(* PLC project station_cds.project, CODESYS CODESYS V3.5 SP22 Patch 1 *)
(* stored: creationDateTime 2026-11-25T17:27:32.309646, modificationDateTime 2026-11-25T17:27:31.3827148 *)

FUNCTION_BLOCK FB_HandleStation
  VAR_INPUT
    CycleTime : REAL := 0.002;  (* s *)
    SafetyOk : BOOL;
    DriveOk : BOOL;
    AckFault : BOOL;
    StartEnable : BOOL;  (* release from the line *)
    PartPresent : BOOL;
    SensLH : BOOL;  (* variant sensor that only an LH unit covers *)
    SensRH : BOOL;  (* variant sensor that only an RH unit covers *)
    VariantLH : BOOL;  (* recipe: TRUE = LH units are being built *)
    ClampClosed : BOOL;
    ClampOpen : BOOL;
    RejectChute : BOOL;  (* light barrier in the reject chute *)
    Pos : REAL;  (* mm, axis position, 0 = home *)
    Force : REAL;  (* N, load cell *)
    VPull : REAL := 50.0;  (* mm/s *)
    VHome : REAL := 150.0;  (* mm/s *)
    FTouch : REAL := 1.5;  (* N *)
    FRev : REAL := 40.0;  (* N *)
    FAbsMax : REAL := 60.0;  (* N, protects the painted part *)
    XMax : REAL := 38.0;  (* mm *)
    TouchLo : REAL := 3.0;  (* mm, window of the touch position *)
    TouchHi : REAL := 7.0;
    Compliance : REAL := 0.025;  (* mm/N, rig deflection taken out of the travel *)
    TareTol : REAL := 0.5;  (* N *)
    TPresent : REAL := 0.1;  (* s *)
    TClampMax : REAL := 1.0;  (* s *)
    TRejectWarn : REAL := 30.0;  (* s *)
    MaxConsecNok : INT := 3;
  END_VAR
  VAR_IN_OUT
    Rcp : ST_EvalRecipe;  (* evaluation recipe, copied into Eval at every tare *)
  END_VAR
  VAR_OUTPUT
    QClamp : BOOL;
    QDriveEnable : BOOL;
    QVel : REAL;  (* mm/s, positive = pull *)
    QLampOk : BOOL;
    QLampNok : BOOL;
    QCallOperator : BOOL;
    State : INT;
    Verdict : INT;  (* 0 none, 1 OK, 2 NOK *)
    NokCode : INT;
    FaultCode : INT;
    Locked : BOOL;
    RigCheckRequired : BOOL;  (* too many rejects in a row: run the master part *)
    XTravel : REAL;  (* mm *)
    FNet : REAL;  (* N *)
    TCycle : REAL;  (* s, clamp to verdict of the last part *)
    CntTotal : DINT;
    CntOk : DINT;
    CntNok : DINT;
    CntRejectConfirmed : DINT;
    CntConsecNok : INT;
    CntByCode : ARRAY[0..31] OF DINT;
  END_VAR
  VAR
    Eval : FB_CurveEval;
    sTim : REAL;
    sTCycle : REAL;
    sTare : REAL;
    sTouchPos : REAL;
    sFTouch : REAL;
    sPreNok : INT;
    sPartGone : BOOL;
    sChutePrev : BOOL;
    sInTest : BOOL;
    sWasLocked : BOOL;
    sState : INT;
    sRigCheckRequired : BOOL;
    sCntTotal : DINT;
    sCntOk : DINT;
    sCntNok : DINT;
    sCntRejectConfirmed : DINT;
    sCntConsecNok : INT;
    sCntByCode : ARRAY[0..31] OF DINT;
  END_VAR
  VAR_TEMP
    tVariantOk : BOOL;
    tChuteEdge : BOOL;
    tCode : INT;
  END_VAR

                {region "Inputs"}
        FNet := Force - sTare;
        tChuteEdge := RejectChute AND NOT sChutePrev;
        sChutePrev := RejectChute;
        sTim := sTim + CycleTime;
        sTCycle := sTCycle + CycleTime;
        QVel := 0.0;
        // exactly the sensor of the expected hand, and not the other one
        tVariantOk := (VariantLH AND SensLH AND NOT SensRH) OR (NOT VariantLH AND SensRH AND NOT SensLH);
    {endregion}

    {region "Faults"}
        IF sState <> 9 AND (NOT SafetyOk OR NOT DriveOk) THEN
            IF NOT SafetyOk THEN
                FaultCode := 1;
            ELSE
                FaultCode := 2;
            END_IF;
            IF sState <> 10 THEN
                sInTest := sState >= 1 AND sState <= 6;
                sWasLocked := sState = 8;
            END_IF;
            sState := 9;
        END_IF;
    {endregion}

    {region "Sequence"}
        CASE sState OF
            0:  // Idle
                Locked := FALSE;
                IF NOT PartPresent THEN
                    sTim := 0.0;
                    QLampOk := FALSE;
                    QLampNok := FALSE;
                ELSIF sTim >= TPresent AND StartEnable AND ClampOpen AND NOT sRigCheckRequired THEN
                    Verdict := 0;
                    NokCode := 0;
                    sPreNok := 0;
                    sTCycle := 0.0;
                    sTim := 0.0;
                    IF tVariantOk THEN
                        sState := 1;
                    ELSE
                        sPreNok := 20;   // never pull a part of the wrong hand
                        sState := 6;
                    END_IF;
                END_IF;
            1:  // Clamp
                QClamp := TRUE;
                IF ClampClosed THEN
                    sTim := 0.0;
                    sState := 2;
                ELSIF sTim > TClampMax THEN
                    FaultCode := 3;
                    sInTest := TRUE;
                    sState := 9;
                END_IF;
            2:  // Tare
                IF sTim >= 0.05 THEN
                    IF ABS(Force) > TareTol THEN
                        FaultCode := 4;
                        sInTest := TRUE;
                        sState := 9;
                    ELSE
                        sTare := Force;
                        // the recipe of this part (Siemens: written into Eval by the caller)
                        Eval.Mode := Rcp.Mode;
                        Eval.GateX := Rcp.GateX;
                        Eval.Gate2X := Rcp.Gate2X;
                        Eval.PeakXLo := Rcp.PeakXLo;
                        Eval.PeakXHi := Rcp.PeakXHi;
                        Eval.StepSpan := Rcp.StepSpan;
                        Eval.StopF := Rcp.StopF;
                        Eval.G1Lo := Rcp.G1Lo;
                        Eval.G1Hi := Rcp.G1Hi;
                        Eval.MeanLo := Rcp.MeanLo;
                        Eval.MeanHi := Rcp.MeanHi;
                        Eval.HystLo := Rcp.HystLo;
                        Eval.HystHi := Rcp.HystHi;
                        Eval.RetFMin := Rcp.RetFMin;
                        Eval.G2Lo := Rcp.G2Lo;
                        Eval.G2Hi := Rcp.G2Hi;
                        Eval.PeakFLo := Rcp.PeakFLo;
                        Eval.PeakFHi := Rcp.PeakFHi;
                        Eval.PeakXMin := Rcp.PeakXMin;
                        Eval.PeakXMax := Rcp.PeakXMax;
                        Eval.StepLo := Rcp.StepLo;
                        Eval.StopXLo := Rcp.StopXLo;
                        Eval.StopXHi := Rcp.StopXHi;
                        Eval.EnvX0 := Rcp.EnvX0;
                        Eval.EnvDx := Rcp.EnvDx;
                        Eval.EnvN := Rcp.EnvN;
                        Eval.EnvLo := Rcp.EnvLo;
                        Eval.EnvHi := Rcp.EnvHi;
                        Eval(Reset := TRUE, Sample := FALSE, Stroke := 0, X := 0.0, F := 0.0, Finish := FALSE);
                        sState := 3;
                    END_IF;
                END_IF;
            3:  // Approach
                QVel := VPull;
                IF FNet > FTouch THEN
                    sTouchPos := Pos;
                    sFTouch := FNet;
                    IF Pos < TouchLo OR Pos > TouchHi THEN
                        sPreNok := 21;
                        sState := 5;
                    ELSE
                        XTravel := 0.0;
                        Eval(Reset := FALSE, Sample := TRUE, Stroke := 1, X := 0.0, F := FNet, Finish := FALSE);
                        sState := 4;
                    END_IF;
                ELSIF Pos > TouchHi THEN
                    sPreNok := 21;
                    sTouchPos := Pos;
                    sFTouch := 0.0;
                    sState := 5;
                END_IF;
            4:  // Pull
                QVel := VPull;
                XTravel := Pos - sTouchPos - (FNet - sFTouch) * Compliance;
                Eval(Reset := FALSE, Sample := TRUE, Stroke := 1, X := XTravel, F := FNet, Finish := FALSE);
                IF FNet >= FAbsMax THEN
                    sPreNok := 22;
                    sState := 5;
                ELSIF FNet >= FRev THEN
                    sState := 5;
                ELSIF XTravel >= XMax THEN
                    sPreNok := 23;
                    sState := 5;
                END_IF;
            5:  // Return
                XTravel := Pos - sTouchPos - (FNet - sFTouch) * Compliance;
                IF Pos > sTouchPos - 0.5 THEN
                    QVel := -VPull;
                    IF sPreNok = 0 THEN
                        Eval(Reset := FALSE, Sample := TRUE, Stroke := 2, X := XTravel, F := FNet, Finish := FALSE);
                    END_IF;
                ELSIF Pos > 0.05 THEN
                    QVel := -VHome;
                ELSE
                    sState := 6;
                END_IF;
            6:  // Evaluate
                IF sPreNok <> 0 THEN
                    tCode := sPreNok;
                ELSE
                    Eval(Reset := FALSE, Sample := FALSE, Stroke := 0, X := 0.0, F := 0.0, Finish := TRUE);
                    tCode := Eval.NokCode;
                END_IF;
                NokCode := tCode;
                TCycle := sTCycle;
                sCntTotal := sCntTotal + 1;
                sCntByCode[tCode] := sCntByCode[tCode] + 1;
                QClamp := FALSE;
                sTim := 0.0;
                IF tCode = 0 THEN
                    Verdict := 1;
                    sCntOk := sCntOk + 1;
                    sCntConsecNok := 0;
                    QLampOk := TRUE;
                    sState := 7;
                ELSE
                    Verdict := 2;
                    sCntNok := sCntNok + 1;
                    sCntConsecNok := sCntConsecNok + 1;
                    QLampNok := TRUE;
                    sPartGone := FALSE;
                    sState := 8;
                END_IF;
            7:  // UnloadOk
                QClamp := FALSE;
                IF NOT PartPresent AND ClampOpen THEN
                    sTim := 0.0;
                    sState := 0;
                END_IF;
            8:  // RejectLock
                QClamp := FALSE;
                Locked := TRUE;
                IF NOT PartPresent THEN
                    sPartGone := TRUE;
                END_IF;
                QCallOperator := sTim > TRejectWarn OR sRigCheckRequired;
                IF sPartGone AND tChuteEdge THEN
                    sCntRejectConfirmed := sCntRejectConfirmed + 1;
                    sRigCheckRequired := sCntConsecNok >= MaxConsecNok;
                    QCallOperator := sRigCheckRequired;
                    Locked := FALSE;
                    sTim := 0.0;
                    sState := 0;
                END_IF;
            9:  // Fault
                QClamp := sInTest;
                QCallOperator := TRUE;
                IF AckFault AND SafetyOk AND DriveOk THEN
                    FaultCode := 0;
                    QCallOperator := FALSE;
                    sState := 10;
                END_IF;
            10:  // Home
                IF Pos > 0.05 THEN
                    QVel := -VPull;
                ELSIF sInTest THEN
                    sInTest := FALSE;
                    sPreNok := 24;
                    sState := 6;
                ELSIF sWasLocked THEN
                    sWasLocked := FALSE;   // a fault does not release the reject lock
                    sState := 8;
                ELSE
                    sState := 0;
                END_IF;
            ELSE
                sState := 9;
        END_CASE;
    {endregion}

    {region "RigCheck"}
        // the lock after too many rejects in a row is released by the acknowledge key
        IF sRigCheckRequired AND AckFault AND sState = 0 THEN
            sRigCheckRequired := FALSE;
            sCntConsecNok := 0;
            QCallOperator := FALSE;
        END_IF;
        QDriveEnable := SafetyOk AND DriveOk AND sState <> 9;
    {endregion}

    {region "Outputs"}
        // state and counters live in static variables; these outputs are written here and nowhere else
        State := sState;
        RigCheckRequired := sRigCheckRequired;
        CntTotal := sCntTotal;
        CntOk := sCntOk;
        CntNok := sCntNok;
        CntRejectConfirmed := sCntRejectConfirmed;
        CntConsecNok := sCntConsecNok;
        CntByCode := sCntByCode;
    {endregion}

          
END_FUNCTION_BLOCK
